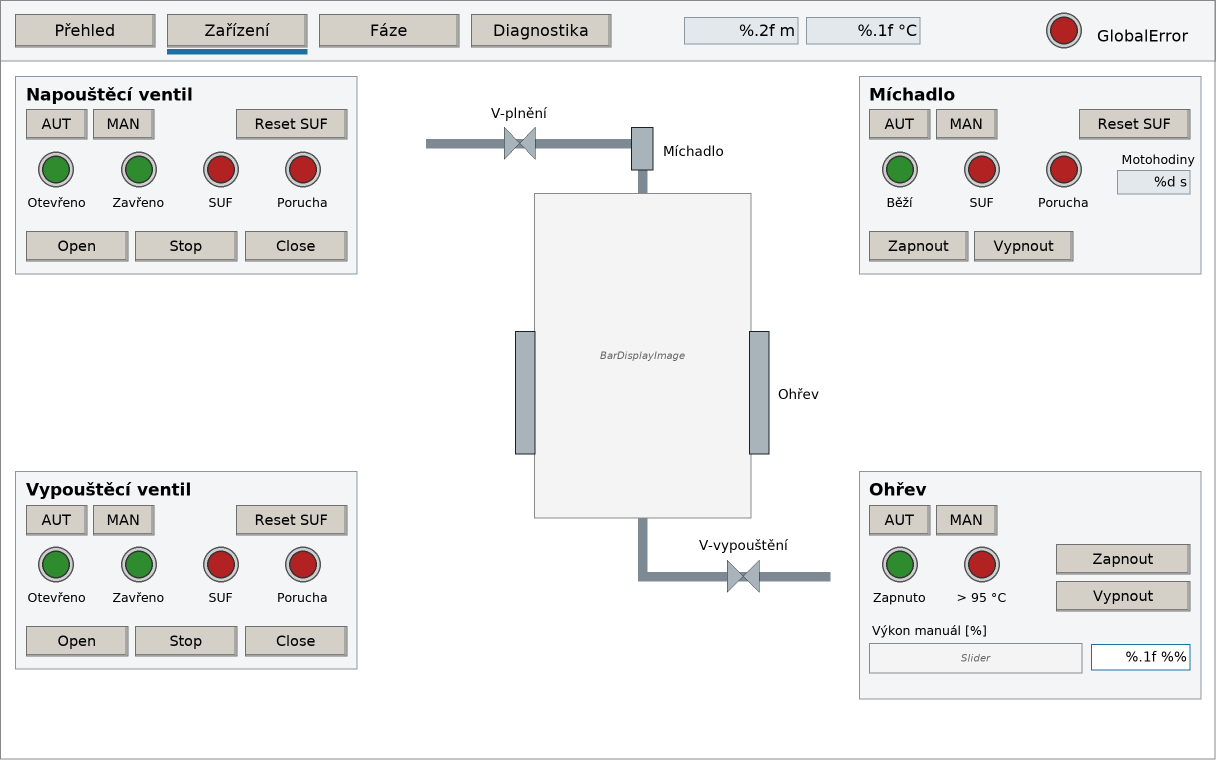
VISUALIZATION Zarizeni  // 1216x760
    Rectangle (0,0 1216x61)
    Button (15,14 140x33), "Přehled"
        OnMouseClick: change screen: Prehled
    Button (167,14 140x33), "Zařízení"
        OnMouseClick: change screen: Zarizeni
    Rectangle (167,49 140x5)
    Button (319,14 140x33), "Fáze"
        OnMouseClick: change screen: Faze
    Button (471,14 140x33), "Diagnostika"
        OnMouseClick: change screen: Diagnostika
    Rectangle (684,17 114x27), "%.2f m", text variable: Global.Tank1.Filling.WaterLevel
    Rectangle (806,17 114x27), "%.1f °C", text variable: Global.Tank1.Heating.WaterTemp
    Lamp1 (1041,10 46x41), variable: Global.Tank1.GlobalError, style: Lamp-Lamp1-Red
    Label (1094,23 126x26), "GlobalError"
    Rectangle (426,139 221x9)
    Rectangle (638,139 9x56)
    Rectangle (638,517 9x64)
    Rectangle (638,572 192x9)
    BarDisplayImage (534,193 217x325), value: Global.Tank1.Filling.WaterLevel, style: BarDisplayImage-Gray, scale format: %.1f, scale 0..2
    Polygon (504,127) (535,159) (535,127) (504,159) (504,159), colour toggle: Global.Tank1.ValveFilling.State.Open
    Label (481,102 76x23), "V-plnění"
    Polygon (727,560) (759,592) (759,560) (727,592) (727,592), colour toggle: Global.Tank1.ValveDraining.State.Open
    Label (698,534 91x23), "V-vypouštění"
    Rectangle (631,127 22x43), colour toggle: Global.Tank1.Mixer.State.Run
    Label (660,140 80x23), "Míchadlo"
    Rectangle (515,331 20x123), colour toggle: Global.Tank1.Heater.State.EnableOut
    Rectangle (749,331 20x123), colour toggle: Global.Tank1.Heater.State.EnableOut
    Label (775,383 52x23), "Ohřev"
    Rectangle (15,76 342x198)
    Label (23,81 201x27), "Napouštěcí ventil"
    Button (26,109 61x30), "AUT", colour toggle: Global.Tank1.ValveFilling.State.AutCtrl
        tap Global.Tank1.ValveFilling.Cmd.AutCtrl
    Button (93,109 61x30), "MAN", colour toggle: Global.Tank1.ValveFilling.State.ManCtrl
        tap Global.Tank1.ValveFilling.Cmd.ManCtrl
    Button (236,109 111x30), "Reset SUF", colour toggle: Global.Tank1.ValveFilling.State.StartupFail
        tap Global.Tank1.ValveFilling.Cmd.ResetSUF
    Lamp1 (33,149 46x41), variable: Global.Tank1.ValveFilling.State.Open, style: Lamp-Lamp1-Green
    Label (11,192 91x21), "Otevřeno"
    Lamp1 (116,149 46x41), variable: Global.Tank1.ValveFilling.State.Closed, style: Lamp-Lamp1-Green
    Label (93,192 91x21), "Zavřeno"
    Lamp1 (198,149 46x41), variable: Global.Tank1.ValveFilling.State.StartupFail, style: Lamp-Lamp1-Red
    Label (175,192 91x21), "SUF"
    Lamp1 (280,149 46x41), variable: Global.Tank1.ValveFilling.State.Err, style: Lamp-Lamp1-Red
    Label (257,192 91x21), "Porucha"
    Button (26,231 102x30), "Open", colour toggle: Global.Tank1.ValveFilling.State.Open
        tap Global.Tank1.ValveFilling.Cmd.OpenMan
    Button (135,231 102x30), "Stop"
        tap Global.Tank1.ValveFilling.Cmd.StopMan
    Button (245,231 102x30), "Close", colour toggle: Global.Tank1.ValveFilling.State.Closed
        tap Global.Tank1.ValveFilling.Cmd.CloseMan
    Rectangle (859,76 342x198)
    Label (866,81 99x27), "Míchadlo"
    Button (869,109 61x30), "AUT", colour toggle: Global.Tank1.Mixer.State.AutCtrl
        tap Global.Tank1.Mixer.Cmd.AutCtrl
    Button (936,109 61x30), "MAN", colour toggle: Global.Tank1.Mixer.State.ManCtrl
        tap Global.Tank1.Mixer.Cmd.ManCtrl
    Button (1079,109 111x30), "Reset SUF", colour toggle: Global.Tank1.Mixer.State.StartUpFail
        tap Global.Tank1.Mixer.Cmd.ResetSUF
    Lamp1 (877,149 46x41), variable: Global.Tank1.Mixer.State.Run, style: Lamp-Lamp1-Green
    Label (854,192 91x21), "Běží"
    Lamp1 (959,149 46x41), variable: Global.Tank1.Mixer.State.StartUpFail, style: Lamp-Lamp1-Red
    Label (936,192 91x21), "SUF"
    Lamp1 (1041,149 46x41), variable: Global.Tank1.Mixer.State.Err, style: Lamp-Lamp1-Red
    Label (1018,192 91x21), "Porucha"
    Button (869,231 99x30), "Zapnout", colour toggle: Global.Tank1.Mixer.State.Run
        tap Global.Tank1.Mixer.Cmd.TurnOnMan
    Button (974,231 99x30), "Vypnout"
        tap Global.Tank1.Mixer.Cmd.TurnOffMan
    Label (1122,149 73x21), "Motohodiny"
    Rectangle (1117,170 73x24), "%d s", text variable: Global.Tank1.Mixer.State.RT
    Rectangle (15,471 342x198)
    Label (23,476 201x27), "Vypouštěcí ventil"
    Button (26,505 61x30), "AUT", colour toggle: Global.Tank1.ValveDraining.State.AutCtrl
        tap Global.Tank1.ValveDraining.Cmd.AutCtrl
    Button (93,505 61x30), "MAN", colour toggle: Global.Tank1.ValveDraining.State.ManCtrl
        tap Global.Tank1.ValveDraining.Cmd.ManCtrl
    Button (236,505 111x30), "Reset SUF", colour toggle: Global.Tank1.ValveDraining.State.StartupFail
        tap Global.Tank1.ValveDraining.Cmd.ResetSUF
    Lamp1 (33,544 46x41), variable: Global.Tank1.ValveDraining.State.Open, style: Lamp-Lamp1-Green
    Label (11,587 91x21), "Otevřeno"
    Lamp1 (116,544 46x41), variable: Global.Tank1.ValveDraining.State.Closed, style: Lamp-Lamp1-Green
    Label (93,587 91x21), "Zavřeno"
    Lamp1 (198,544 46x41), variable: Global.Tank1.ValveDraining.State.StartupFail, style: Lamp-Lamp1-Red
    Label (175,587 91x21), "SUF"
    Lamp1 (280,544 46x41), variable: Global.Tank1.ValveDraining.State.Err, style: Lamp-Lamp1-Red
    Label (257,587 91x21), "Porucha"
    Button (26,626 102x30), "Open", colour toggle: Global.Tank1.ValveDraining.State.Open
        tap Global.Tank1.ValveDraining.Cmd.OpenMan
    Button (135,626 102x30), "Stop"
        tap Global.Tank1.ValveDraining.Cmd.StopMan
    Button (245,626 102x30), "Close", colour toggle: Global.Tank1.ValveDraining.State.Closed
        tap Global.Tank1.ValveDraining.Cmd.CloseMan
    Rectangle (859,471 342x228)
    Label (866,476 65x27), "Ohřev"
    Button (869,505 61x30), "AUT", colour toggle: Global.Tank1.Heater.State.AutCtrl
        tap Global.Tank1.Heater.Cmd.AutCtrl
    Button (936,505 61x30), "MAN", colour toggle: Global.Tank1.Heater.State.ManCtrl
        tap Global.Tank1.Heater.Cmd.ManCtrl
    Lamp1 (877,544 46x41), variable: Global.Tank1.Heater.State.EnableOut, style: Lamp-Lamp1-Green
    Label (854,587 91x21), "Zapnuto"
    Lamp1 (959,544 46x41), variable: Global.Tank1.Heater.State.GenErr, style: Lamp-Lamp1-Red
    Label (936,587 91x21), "> 95 °C"
    Button (1056,544 134x30), "Zapnout", colour toggle: Global.Tank1.Heater.State.EnableOut
        tap Global.Tank1.Heater.Cmd.TurnOnMan
    Button (1056,581 134x30), "Vypnout"
        tap Global.Tank1.Heater.Cmd.TurnOffMan
    Label (869,620 142x21), "Výkon manuál [%]"
    Slider (869,643 213x30), variable: Global.Tank1.Heater.ParamHeatingPowerManual, scale 0..100
    Rectangle (1091,644 99x26), "%.1f %%", text variable: Global.Tank1.Heater.ParamHeatingPowerManual
        OnMouseClick: write the text variable via Default
END_VISUALIZATION

(* stored: Version 1.1.0.1, ProductVersion 3.1.4024.16
   Visu Zarizeni: Id {fb3cfcc8-39d1-482d-9945-8cc44f70ca12} *)
